(* IEC 61131-3 sources: PLC-Static-Analysis/modules/plc-semantic/src/test/resources/dev/plca/semantic/SemanticFuzzTestInputs/fuzzModel, 6 files *)

(* ---- types.st ---- *)
{attribute 'qualified_only'}
{attribute 'strict'}
TYPE E_State : (Idle, Starting := 5, Running, Faulted) INT;
END_TYPE

TYPE E_Mode : (Manual, Auto);
END_TYPE

TYPE
    ST_Base :
    STRUCT
        nId : UDINT;
    END_STRUCT
    ST_Motor EXTENDS ST_Base :
    STRUCT
        rSpeed : REAL;
        aLog : ARRAY[0..LOG_SIZE - 1] OF INT;
    END_STRUCT
    T_Speed : REAL;
END_TYPE

(* ---- GVL_Main.st ---- *)
VAR_GLOBAL CONSTANT
    LOG_SIZE : INT := 10;
END_VAR
VAR_GLOBAL
    gnCounter : DINT;
    gAxis : Tc2_MC2.AXIS_REF;
END_VAR

(* ---- functions.st ---- *)
FUNCTION F_Scale : REAL
VAR_INPUT
    rIn : REAL;
    nDepth : INT;
END_VAR
IF nDepth > 0 THEN
    F_Scale := F_Helper(rIn, nDepth - 1);
ELSE
    F_Scale := rIn * 2.5;
END_IF
END_FUNCTION

FUNCTION F_Helper : REAL
VAR_INPUT
    rIn : REAL;
    nDepth : INT;
END_VAR
F_Helper := F_Scale(rIn := rIn, nDepth := nDepth);
END_FUNCTION

(* ---- FB_Base.st ---- *)
FUNCTION_BLOCK ABSTRACT FB_Base
VAR_INPUT
    bEnable : BOOL;
END_VAR
VAR
    nCalls : INT;
END_VAR
nCalls := nCalls + 1;

METHOD PUBLIC Reset : BOOL
nCalls := 0;
Reset := TRUE;
END_METHOD
END_FUNCTION_BLOCK

(* ---- FB_Motor.st ---- *)
FUNCTION_BLOCK FB_Motor EXTENDS FB_Base
VAR_INPUT
    rSetpoint : T_Speed;
END_VAR
VAR_OUTPUT
    bRunning : BOOL;
END_VAR
VAR_IN_OUT
    stData : ST_Motor;
END_VAR
VAR
    fbDelay : Tc2_Standard.TON;
    fbPower : Tc2_MC2.MC_Power;
    eState : E_State;
    pData : POINTER TO ST_Motor;
END_VAR

fbDelay(IN := bEnable, PT := T#500MS, Q => bRunning);
CASE eState OF
    Idle: IF bEnable THEN eState := E_State.Starting; END_IF
    Starting: eState := E_State.Running;
END_CASE
stData.aLog[3] := nCalls;
stData.rSpeed := rSetpoint;
pData := ADR(stData);
fbPower(Axis := gAxis, Enable := bEnable);
Stop();

METHOD PUBLIC Reset : BOOL
bRunning := FALSE;
Reset := SUPER^.Reset();
END_METHOD

PROPERTY PUBLIC Speed : REAL
GET
    Speed := stData.rSpeed;
END_GET
END_PROPERTY

ACTION Stop:
    bRunning := FALSE;
END_ACTION
END_FUNCTION_BLOCK

(* ---- MAIN.st ---- *)
PROGRAM MAIN
VAR
    fbMotor : FB_Motor;
    aMotors : ARRAY[1..2] OF FB_Motor;
    stMotor : ST_Motor;
    rSpeed : REAL;
    n : DINT;
    i : INT;
    eMode : E_Mode;
END_VAR
fbMotor(bEnable := GVL_IO.bStart, rSetpoint := 1500.0, stData := stMotor);
rSpeed := fbMotor.Speed + F_Scale(rSpeed, 3);
n := i + 1;
FOR i := 1 TO 2 DO
    aMotors[i](stData := stMotor);
END_FOR
gnCounter := gnCounter + 1;
eMode := Auto;
IF fbMotor.Reset() THEN
    ;
END_IF
END_PROGRAM

PROGRAM FAST
gnCounter := 0;
END_PROGRAM
